TYPE ST_EVENT : 
STRUCT
	eEventType : Tc2_System.TcEvent;
	eEventSeverity : Global.TcEventSeverity;
	nEventIdentity : UDINT;
	sEventText : STRING(255);
	dtTimeStamp : DATE_AND_TIME;
END_STRUCT
END_TYPE

(* stored: Version 1.1.0.1
   DUT ST_EVENT: Id {e290a143-334c-4540-9367-c877fa98893d} *)
